// Where the transport orders come from.
{attribute 'qualified_only'}
{attribute 'strict'}
TYPE E_MfrLink :
(
    eEmulator := 0,   // FB_MfrEmulator in the PLC (commissioning, demo, tests)
    eTcp      := 1    // real material flow computer over TCP/IP (PLC is the server)
) INT;
END_TYPE

(* stored: Version 1.1.0.1
   DUT E_MfrLink: Id {51bd9ef0-a111-b88e-c483-6405f97fa508} *)
